Fanuc KAREL source: ko00055.KL

-- PROVISIONAL review KL for V1013-1; original PC SHA256 1b0802369a168d54738684c532b970294376e26cb5d55af2253e0bc19f8b92be
-- Incomplete behavior may be omitted. Consult companion uncertainty JSON. Do not deploy.
PROGRAM KO00055
%NOLOCKGROUP
BEGIN
  -- UNRESOLVED_PC offsets 5-12; opcodes 9D,23
  -- UNRESOLVED_PC offsets 17-69; opcodes 27,27,49,7E,AD,27,49,7E,AD,22,31,7E,4A
  -- UNRESOLVED_PC offsets 74-78; opcodes 7F
END KO00055
